# EPICS autosave request: iocs/meascomp/db/measCompTemperatureIn_settings.req
$(P)$(R)Scale
$(P)$(R)TCType
$(P)$(R)OpenTCDetect
$(P)$(R)Filter
$(P)$(R).LOPR
$(P)$(R).HOPR
$(P)$(R).PREC
$(P)$(R).SCAN
